Fanuc KAREL source: kf00046.KL

-- PROVISIONAL review KL for V1013-1; original PC SHA256 dc8ebb778b904a0c91eace24575742de9a1cbe94f4a1ca6869e071ea5e341dd5
-- Incomplete behavior may be omitted. Consult companion uncertainty JSON. Do not deploy.
PROGRAM KF00046
%NOLOCKGROUP
VAR
  I : INTEGER
  J : INTEGER
  X : REAL
  Y : REAL
  B : BOOLEAN
  C : BOOLEAN
  TXT : STRING[80]
  TXT2 : STRING[80]
  STATUS : INTEGER
-- UNRESOLVED_DECL AI type=002010
-- UNRESOLVED_DECL BI type=002010
-- UNRESOLVED_DECL P type=000102
-- UNRESOLVED_DECL JP type=000199
-- UNRESOLVED_DECL PF type=000101
-- UNRESOLVED_DECL V1 type=000013
-- UNRESOLVED_DECL V2 type=000013
BEGIN
  -- UNRESOLVED_PC offsets 5-12; opcodes 9D,23
  -- UNRESOLVED_PC offsets 17-30; opcodes 21,9D,57,79
  -- UNRESOLVED_PC offsets 35-46; opcodes 2E,23
  -- UNRESOLVED_PC offsets 51-56; opcodes 7A
  -- UNRESOLVED_PC offsets 61-72; opcodes 2E,23
  -- UNRESOLVED_PC offsets 82-86; opcodes 7F
END KF00046
